// TIA Portal V21 export
// export: Created 2026-10-12T11:32:14.1584136Z, ExportSetting WithDefaults, DisplayName Totally Integrated Automation Portal, DisplayVersion V21, DisplayName STEP 7 Professional, DisplayVersion V21, DisplayName STEP 7 Safety, DisplayVersion V21, DisplayName Tech WebApplication, DisplayVersion V21, DisplayName WinCC Basic/Comfort/Advanced, DisplayVersion V21, DisplayName WinCC Unified, DisplayVersion V21
FUNCTION "FC_ALARMS" : Void   // FC3, LAD
{ S7_Optimized_Access := 'TRUE' }
VERSION : 0.1
// stored: AutoNumber true, IsIECCheckEnabled false, SetENOAutomatically false, UDAEnableTagReadback false
BEGIN

REGION Network 1: EMERGENCY PB PRESSED FAULT (I0.4)
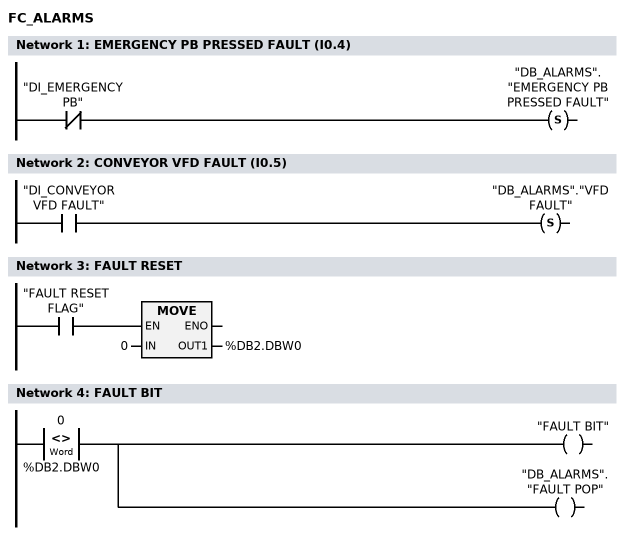
   RUNG wire#powerrail
      I_Contact( "DI_EMERGENCY PB" )
      S_Coil( "DB_ALARMS"."EMERGENCY PB PRESSED FAULT" )
   END_RUNG
   // the same network as SCL:
   IF NOT "DI_EMERGENCY PB" THEN "DB_ALARMS"."EMERGENCY PB PRESSED FAULT" := TRUE; END_IF;
END_REGION

REGION Network 2: CONVEYOR VFD FAULT (I0.5)
   RUNG wire#powerrail
      Contact( "DI_CONVEYOR VFD FAULT" )
      S_Coil( "DB_ALARMS"."VFD FAULT" )
   END_RUNG
   // the same network as SCL:
   IF "DI_CONVEYOR VFD FAULT" THEN "DB_ALARMS"."VFD FAULT" := TRUE; END_IF;
END_REGION

REGION Network 3: FAULT RESET
   RUNG wire#powerrail
      Contact( "FAULT RESET FLAG" )
      Move(in := 0, out1 => %DB2.DBW0)
   END_RUNG
   // the same network as SCL:
   IF "FAULT RESET FLAG" THEN %DB2.DBW0 := 0; END_IF;
END_REGION

REGION Network 4: FAULT BIT
   RUNG wire#powerrail
      { S7_Templates := "SrcType := Word" } NE_Contact(in1 := 0, in2 := %DB2.DBW0)
      wire#w1
      Coil( "FAULT BIT" )
   END_RUNG
   RUNG wire#w1
      Coil( "DB_ALARMS"."FAULT POP" )
   END_RUNG
   // the same network as SCL:
   "FAULT BIT" := 0 <> %DB2.DBW0;
   "DB_ALARMS"."FAULT POP" := "FAULT BIT";
END_REGION
END_FUNCTION
